// TIA Portal V20 export
// export: Created 2026-10-06T00:00:00
Screen "Conveyor_Overview"  1280x800, Number=2, Template=Base
  ScreenLayer 
    Rectangle "Motor_1" at 60,100 size 40x40
      VisibilityAnimation "VisibilityAnimation"
        tag Motor_1_Run
